Yaskawa INFORM job: 20211127CHUFENGKOUSAVE.JBI

/JOB
//NAME 20211127CHUFENGKOUSAVE
//POS
///NPOS 7,0,7,0,0,0
///TOOL 1
///POSTYPE PULSE
///PULSE
C00000=-5456,29378,14097,-3416,-76919,3294
C00001=-5457,32223,-10944,-3917,-57557,3928
C00002=-5334,32532,-16573,-4115,-53450,4056
C00003=-5334,32532,-16573,-4115,-53450,4056
C00004=-5335,32532,-16573,-4114,-53450,4057
C00005=-5253,34423,-13635,-4085,-54045,4006
C00006=-5387,38273,25473,-3407,-78050,3239
///TOOL 0
EC00000=-4,321083
EC00001=-4,321083
EC00002=-4,321083
EC00003=-4,321083
EC00004=-4,221835
EC00005=-4,93195
EC00006=-4,93198
//INST
///DATE 2021/11/27 11:12
///ATTR SC,RW
///GROUP1 RB1
///GROUP2 ST1
NOP
MOVJ C00000 VJ=10.00  +MOVJ EC00000 VJ=10.00
MOVJ C00001 VJ=10.00  +MOVJ EC00001 VJ=0.78
MOVL C00002 V=20.0  +MOVJ EC00002 VJ=10.00
CALL JOB:SAVETRAJ
SMOVC C00003 V=20.0  +MOVJ EC00003
SMOVC C00004 V=4.5  +MOVJ EC00004
SMOVC C00005 V=4.5  +MOVJ EC00005
MOVL C00006 V=20.0  +MOVJ EC00006 VJ=10.00
END
